(* IEC 61131-3 sources: llm-plc-st-eval/data/processed_definitivo/claude-sonnet-4-6/I2/zero_shot, 3 files *)

(* ---- ejec_1.st ---- *)
FUNCTION_BLOCK FB_Llenado
VAR_INPUT
    nivelAlto  : BOOL; (* Sensor de nivel alto *)
    nivelBajo  : BOOL; (* Sensor de nivel bajo *)
    btnInicio  : BOOL; (* Botón de inicio (flanco) *)
    btnParo    : BOOL; (* Botón de paro (nivel) *)
END_VAR

VAR_OUTPUT
    vLlenado    : BOOL; (* Válvula de llenado *)
    motorMezcla : BOOL; (* Motor de mezcla *)
    vDescarga   : BOOL; (* Válvula de descarga *)
END_VAR

VAR
    (* Etapas del proceso *)
    eEtapa : INT := 0;
    (*
        0 = Reposo
        1 = Llenado
        2 = Mezcla
        3 = Descarga
    *)

    (* Temporizador para la etapa de mezcla *)
    tonMezcla : TON;

    (* Detección de flanco ascendente en btnInicio *)
    rTrigInicio : R_TRIG;
END_VAR

(* ─────────────────────────────────────────────
   Detección de flanco ascendente en btnInicio
   ───────────────────────────────────────────── *)
rTrigInicio(CLK := btnInicio);

(* ─────────────────────────────────────────────
   Paro de emergencia: cualquier etapa
   ───────────────────────────────────────────── *)
IF btnParo THEN
    eEtapa      := 0;
    vLlenado    := FALSE;
    motorMezcla := FALSE;
    vDescarga   := FALSE;
    tonMezcla(IN := FALSE, PT := T#60S); (* Resetea temporizador *)
    RETURN; (* Sale del bloque sin ejecutar el resto *)
END_IF;

(* ─────────────────────────────────────────────
   Máquina de estados
   ───────────────────────────────────────────── *)
CASE eEtapa OF

    (* ── Etapa 0: Reposo ── *)
    0:
        vLlenado    := FALSE;
        motorMezcla := FALSE;
        vDescarga   := FALSE;
        tonMezcla(IN := FALSE, PT := T#60S); (* Mantiene temporizador reseteado *)

        IF rTrigInicio.Q THEN
            eEtapa := 1; (* Ir a llenado *)
        END_IF;

    (* ── Etapa 1: Llenado ── *)
    1:
        vLlenado    := TRUE;
        motorMezcla := FALSE;
        vDescarga   := FALSE;

        IF nivelAlto THEN
            vLlenado := FALSE;
            eEtapa   := 2; (* Ir a mezcla *)
        END_IF;

    (* ── Etapa 2: Mezcla (60 s) ── *)
    2:
        vLlenado    := FALSE;
        motorMezcla := TRUE;
        vDescarga   := FALSE;
        tonMezcla(IN := TRUE, PT := T#60S); (* Arranca/mantiene temporizador *)

        IF tonMezcla.Q THEN
            motorMezcla := FALSE;
            tonMezcla(IN := FALSE, PT := T#60S); (* Resetea para próximo ciclo *)
            eEtapa := 3; (* Ir a descarga *)
        END_IF;

    (* ── Etapa 3: Descarga ── *)
    3:
        vLlenado    := FALSE;
        motorMezcla := FALSE;
        vDescarga   := TRUE;

        IF nivelBajo THEN
            vDescarga := FALSE;
            eEtapa    := 0; (* Volver a reposo *)
        END_IF;

    (* ── Estado no definido: seguridad ── *)
    ELSE:
        eEtapa      := 0;
        vLlenado    := FALSE;
        motorMezcla := FALSE;
        vDescarga   := FALSE;

END_CASE;

(* ---- ejec_2.st ---- *)
FUNCTION_BLOCK FB_Llenado
VAR_INPUT
    nivelAlto  : BOOL; (* Sensor de nivel alto *)
    nivelBajo  : BOOL; (* Sensor de nivel bajo *)
    btnInicio  : BOOL; (* Botón de inicio del proceso *)
    btnParo    : BOOL; (* Botón de paro de emergencia *)
END_VAR

VAR_OUTPUT
    vLlenado    : BOOL; (* Válvula de llenado *)
    motorMezcla : BOOL; (* Motor de mezcla *)
    vDescarga   : BOOL; (* Válvula de descarga *)
END_VAR

VAR
    (* Etapas del proceso *)
    eEtapa : INT := 0;
    (*
        0 = Reposo
        1 = Llenado
        2 = Mezcla
        3 = Descarga
    *)

    (* Temporizador para la etapa de mezcla *)
    tonMezcla : TON;
END_VAR

(* ─────────────────────────────────────────────
   Lógica principal
   ───────────────────────────────────────────── *)

(* Paro de emergencia: tiene prioridad sobre cualquier etapa *)
IF btnParo THEN
    eEtapa      := 0;
    vLlenado    := FALSE;
    motorMezcla := FALSE;
    vDescarga   := FALSE;
    tonMezcla(IN := FALSE, PT := T#60S); (* Reinicia temporizador *)

ELSE

    CASE eEtapa OF

        (* ── Etapa 0: Reposo ── *)
        0:
            vLlenado    := FALSE;
            motorMezcla := FALSE;
            vDescarga   := FALSE;
            tonMezcla(IN := FALSE, PT := T#60S);

            IF btnInicio THEN
                eEtapa := 1; (* Ir a llenado *)
            END_IF;

        (* ── Etapa 1: Llenado ── *)
        1:
            vLlenado    := TRUE;
            motorMezcla := FALSE;
            vDescarga   := FALSE;

            IF nivelAlto THEN
                vLlenado := FALSE;
                eEtapa   := 2; (* Ir a mezcla *)
            END_IF;

        (* ── Etapa 2: Mezcla (60 s) ── *)
        2:
            vLlenado    := FALSE;
            motorMezcla := TRUE;
            vDescarga   := FALSE;

            (* Activa el temporizador mientras se está en esta etapa *)
            tonMezcla(IN := TRUE, PT := T#60S);

            IF tonMezcla.Q THEN
                motorMezcla := FALSE;
                tonMezcla(IN := FALSE, PT := T#60S); (* Reinicia para próximo ciclo *)
                eEtapa := 3; (* Ir a descarga *)
            END_IF;

        (* ── Etapa 3: Descarga ── *)
        3:
            vLlenado    := FALSE;
            motorMezcla := FALSE;
            vDescarga   := TRUE;

            IF nivelBajo THEN
                vDescarga := FALSE;
                eEtapa    := 0; (* Volver a reposo *)
            END_IF;

        (* ── Estado no definido: ir a reposo de forma segura ── *)
        ELSE
            eEtapa      := 0;
            vLlenado    := FALSE;
            motorMezcla := FALSE;
            vDescarga   := FALSE;

    END_CASE;

END_IF;

(* ---- ejec_3.st ---- *)
FUNCTION_BLOCK FB_Llenado
VAR_INPUT
    nivelAlto  : BOOL; (* Sensor de nivel alto *)
    nivelBajo  : BOOL; (* Sensor de nivel bajo *)
    btnInicio  : BOOL; (* Botón de inicio del proceso *)
    btnParo    : BOOL; (* Botón de paro de emergencia *)
END_VAR

VAR_OUTPUT
    vLlenado    : BOOL; (* Válvula de llenado *)
    motorMezcla : BOOL; (* Motor de mezcla *)
    vDescarga   : BOOL; (* Válvula de descarga *)
END_VAR

VAR
    etapa       : INT;          (* Etapa actual del proceso: 0=Reposo, 1=Llenado, 2=Mezcla, 3=Descarga *)
    timerMezcla : TON;          (* Temporizador para la etapa de mezcla *)
END_VAR

(* ─────────────────────────────────────────────
   Máquina de estados del proceso de llenado
   ───────────────────────────────────────────── *)

(* Paro de emergencia: actúa en cualquier etapa *)
IF btnParo THEN
    etapa       := 0;
    vLlenado    := FALSE;
    motorMezcla := FALSE;
    vDescarga   := FALSE;
    timerMezcla(IN := FALSE, PT := T#60S); (* Resetea el temporizador *)
ELSE

    CASE etapa OF

        (* ── ETAPA 0: Reposo ── *)
        0:
            vLlenado    := FALSE;
            motorMezcla := FALSE;
            vDescarga   := FALSE;
            timerMezcla(IN := FALSE, PT := T#60S); (* Mantiene timer reseteado *)

            IF btnInicio THEN
                etapa := 1; (* Transición a llenado *)
            END_IF;

        (* ── ETAPA 1: Llenado ── *)
        1:
            vLlenado    := TRUE;
            motorMezcla := FALSE;
            vDescarga   := FALSE;

            IF nivelAlto THEN
                vLlenado := FALSE;
                etapa    := 2; (* Transición a mezcla *)
            END_IF;

        (* ── ETAPA 2: Mezcla (60 segundos) ── *)
        2:
            vLlenado    := FALSE;
            motorMezcla := TRUE;
            vDescarga   := FALSE;

            timerMezcla(IN := TRUE, PT := T#60S); (* Activa el temporizador *)

            IF timerMezcla.Q THEN
                motorMezcla := FALSE;
                timerMezcla(IN := FALSE, PT := T#60S); (* Resetea para próximo ciclo *)
                etapa := 3; (* Transición a descarga *)
            END_IF;

        (* ── ETAPA 3: Descarga ── *)
        3:
            vLlenado    := FALSE;
            motorMezcla := FALSE;
            vDescarga   := TRUE;

            IF nivelBajo THEN
                vDescarga := FALSE;
                etapa     := 0; (* Regresa a reposo *)
            END_IF;

        (* ── Estado no definido: regreso seguro a reposo ── *)
        ELSE
            etapa       := 0;
            vLlenado    := FALSE;
            motorMezcla := FALSE;
            vDescarga   := FALSE;

    END_CASE;

END_IF;
